Fanuc KAREL source: KT00467.KL

PROGRAM KT00467
%NOLOCKGROUP
VAR
  P1: JOINTPOS
  P2: POSITION
  OUT: BOOLEAN
BEGIN
  OUT = P1 >= P2
END KT00467
